Staubli VAL3: MutliMatrix.pgx

public program MutliMatrix(num& x_nMatrix1[] (dimensions=2), num& x_nMatrix2[] (dimensions=2), num& x_nMatrix3[] (dimensions=2))
  local num a11
  local num a12
  local num a13
  local num a14
  local num a21
  local num a22
  local num a23
  local num a24
  local num a31
  local num a32
  local num a33
  local num a34
  local num a41
  local num a42
  local num a43
  local num a44
  local num b11
  local num b12
  local num b13
  local num b14
  local num b21
  local num b22
  local num b23
  local num b24
  local num b31
  local num b32
  local num b33
  local num b34
  local num b41
  local num b42
  local num b43
  local num b44
begin
  //初始化变量
  a11=x_nMatrix1[0,0]
  a21=x_nMatrix1[0,1]
  a31=x_nMatrix1[0,2]
  a41=x_nMatrix1[0,3]
  a12=x_nMatrix1[1,0]
  a22=x_nMatrix1[1,1]
  a32=x_nMatrix1[1,2]
  a42=x_nMatrix1[1,3]
  a13=x_nMatrix1[2,0]
  a23=x_nMatrix1[2,1]
  a33=x_nMatrix1[2,2]
  a43=x_nMatrix1[2,3]
  a14=x_nMatrix1[3,0]
  a24=x_nMatrix1[3,1]
  a34=x_nMatrix1[3,2]
  a44=x_nMatrix1[3,3]

  b11=x_nMatrix2[0,0]
  b21=x_nMatrix2[0,1]
  b31=x_nMatrix2[0,2]
  b41=x_nMatrix2[0,3]
  b12=x_nMatrix2[1,0]
  b22=x_nMatrix2[1,1]
  b32=x_nMatrix2[1,2]
  b42=x_nMatrix2[1,3]
  b13=x_nMatrix2[2,0]
  b23=x_nMatrix2[2,1]
  b33=x_nMatrix2[2,2]
  b43=x_nMatrix2[2,3]
  b14=x_nMatrix2[3,0]
  b24=x_nMatrix2[3,1]
  b34=x_nMatrix2[3,2]
  b44=x_nMatrix2[3,3]

  //矩阵相乘

  x_nMatrix3[0,0]=a11*b11+a12*b21+a13*b31+a14*b41
  x_nMatrix3[0,1]=a21*b11+a22*b21+a23*b31+a24*b41
  x_nMatrix3[0,2]=a31*b11+a32*b21+a33*b31+a34*b41
  x_nMatrix3[0,3]=a41*b11+a42*b21+a43*b31+a44*b41

  x_nMatrix3[1,0]=a11*b12+a12*b22+a13*b32+a14*b42
  x_nMatrix3[1,1]=a21*b12+a22*b22+a23*b32+a24*b42
  x_nMatrix3[1,2]=a31*b12+a32*b22+a33*b32+a34*b42
  x_nMatrix3[1,3]=a41*b12+a42*b22+a43*b32+a44*b42

  x_nMatrix3[2,0]=a11*b13+a12*b23+a13*b33+a14*b43
  x_nMatrix3[2,1]=a21*b13+a22*b23+a23*b33+a24*b43
  x_nMatrix3[2,2]=a31*b13+a32*b23+a33*b33+a34*b43
  x_nMatrix3[2,3]=a41*b13+a42*b23+a43*b33+a44*b43

  x_nMatrix3[3,0]=a11*b14+a12*b24+a13*b34+a14*b44
  x_nMatrix3[3,1]=a21*b14+a22*b24+a23*b34+a24*b44
  x_nMatrix3[3,2]=a31*b14+a32*b24+a33*b34+a34*b44
  x_nMatrix3[3,3]=a41*b14+a42*b24+a43*b34+a44*b44
end
